ABB RobotStudio station: Project2_1.rsstnx

Station Project2 (saved by RobotStudio 25.5.11605.0)
Controller Controller1
  mechanical unit ROB_1: IRB1090_3_58__02, 6 joints, base frame (0, 0, 0) mm
Layout (positions relative to the parent item):
  - IRB1090_3_58__02 [mechanism, from %ABB.RobotStudio.Models.IRB1090%\IRB1090_3_58__01.rslib] at (0, 0, 0) mm; joint values [-0.1802, 0.1972, 0.0337, -0.0141, 1.3827, 4.496] (rad or m)
  - SOURCE AREA [graphiccomponentgroup, from Equipment\Euro Pallet.rslib] at (-200, 120, 0) mm
    - Body 1 [part, from Equipment\Euro Pallet.rslib]
  - RED_SORT_AREA [graphiccomponentgroup, from Equipment\Euro Pallet.rslib] at (-200, -920, 0) mm
    - Body 1 [part, from Equipment\Euro Pallet.rslib]
  - Source_R04 [part], size 150 x 149.2 x 50 mm
  - Source_R02 [part] at (-160, 0, 0) mm, size 150 x 149.2 x 50 mm
  - Source_R05 [part] at (-90, 150, 0) mm, size 150 x 149.2 x 50 mm
  - Source_G04 [part] at (0, 0, 50) mm, size 150 x 149.2 x 50 mm
  - Source_R03 [part] at (0, 0, 100) mm, size 150 x 149.2 x 50 mm
  - Source_G03 [part] at (0, 0, 150) mm, size 150 x 149.2 x 50 mm
  - Source_G02 [part] at (-160, 0, 50) mm, size 150 x 149.2 x 50 mm
  - Source_G01 [part] at (-160, 0, 100) mm, size 150 x 149.2 x 50 mm
  - Source_R01 [part] at (-160, 0, 150) mm, size 150 x 149.2 x 50 mm
  - Source_G07 [part] at (-90, 150, 50) mm, size 150 x 149.2 x 50 mm
  - Source_G06 [part] at (-90, 150, 100) mm, size 150 x 149.2 x 50 mm
  - Source_G05 [part] at (-90, 150, 150) mm, size 150 x 149.2 x 50 mm
  - SG_EE [smart component] at (327.71, -364.56, -73.2) mm, rotated rx 2.57 ry 0.1 rz 92.24 deg
      signals: DI To_Grasp, DO Red_Detected, DO Green_Detected
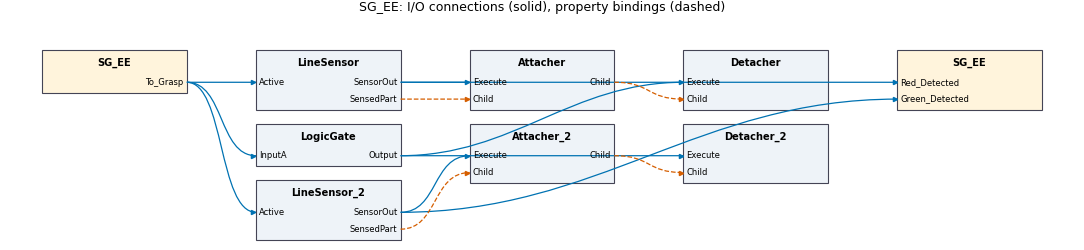
      connections:
        SG_EE.To_Grasp -> LineSensor.Active
        SG_EE.To_Grasp -> LogicGate.InputA
        LogicGate.Output -> Detacher.Execute
        LineSensor.SensorOut -> Attacher.Execute
        SG_EE.To_Grasp -> LineSensor_2.Active
        LineSensor_2.SensorOut -> Attacher_2.Execute
        LogicGate.Output -> Detacher_2.Execute
        LineSensor.SensorOut -> SG_EE.Red_Detected
        LineSensor_2.SensorOut -> SG_EE.Green_Detected
        LineSensor.SensedPart => Attacher.Child
        Attacher.Child => Detacher.Child
        LineSensor_2.SensedPart => Attacher_2.Child
        Attacher_2.Child => Detacher_2.Child
    - LogicGate [smart component, from Components\LogicGate.rslib]
        properties: Operator=NOT; Delay=0
    - LineSensor [smart component, from Components\LineSensor.rslib] at (0, 0, 50) mm
        properties: Start=[0.3 0 0.435]; End=[0.3 0 0.425]; Length=0.00999999999999995; Radius=0.0110132158590308; Tag=Tag_1; SenseMultiple=false; SensedPart=(none); SensedPoint=[0 0 0]
      - _sensorPart_ [part], size 22 x 22 x 10 mm
    - Attacher [smart component, from Components\Attacher.rslib]
        properties: Parent=EE_tool; Flange=0; Child=(none); Mount=false; Offset=[0 0 0]; Orientation=[0 0 0]
    - Detacher [smart component, from Components\Detacher.rslib]
        properties: Child=(none); KeepPosition=true
    - EE_tool [mechanism] at (299.85, 0, 553) mm, rotated rx 180 ry -0.14 rz 180 deg
        TCP EE_tool at (0, 0, -70) mm, rotated rx 180 ry 0 rz 0 deg
        links: EE
    - LineSensor_2 [smart component, from Components\LineSensor.rslib]
        properties: Start=[0.300468401861399 -2.79720985579823E-06 0.484511357513637]; End=[0.300525732933959 0.000547750941646302 0.474476736948762]; Length=0.0100498756211209; Radius=0.0108695652173913; Tag=Tag_2; SenseMultiple=false; SensedPart=(none); SensedPoint=[0 0 0]
      - _sensorPart_ [part], size 21.7 x 22.1 x 11.2 mm
    - Attacher_2 [smart component, from Components\Attacher.rslib]
        properties: Parent=EE_tool; Flange=0; Child=(none); Mount=false; Offset=[0 0 0]; Orientation=[0 0 0]
    - Detacher_2 [smart component, from Components\Detacher.rslib]
        properties: Child=(none); KeepPosition=true
Attachment: EE_tool is attached to IRB1090_3_58__02 / Link6
Attachment: SG_EE is attached to IRB1090_3_58__02 / Link6
Station logic (signal -> signal, property => property):
  Controller1.to_grasp_signal -> SG_EE.To_Grasp
  SG_EE.Red_Detected -> Controller1.red_detect
  SG_EE.Green_Detected -> Controller1.green_detect
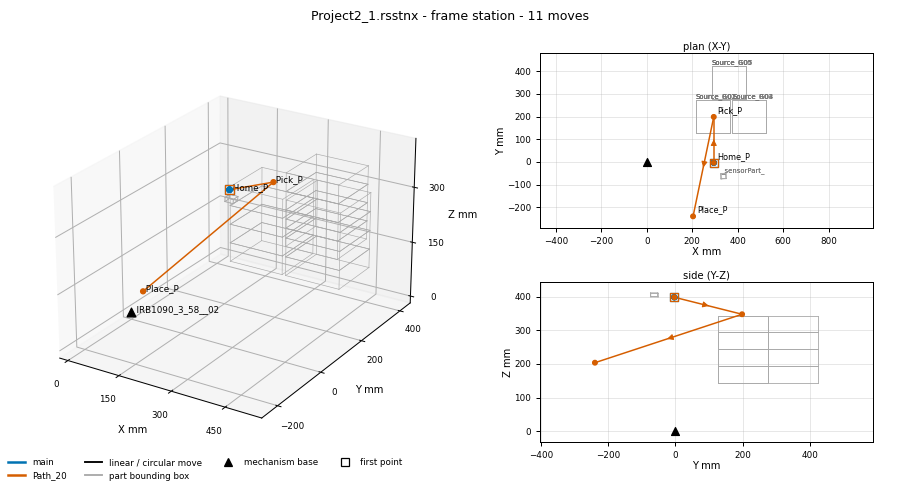
[picture p0: tool path of Project2_1.rsstnx in frame station, 11 of 26 moves have a stored position in this frame; points joined in program order, loops and branches not executed]
Targets, tools, work objects and paths stored in the station, written as RAPID:
! task T_ROB1
MODULE CalibData
  PERS tooldata EE_tool:=[TRUE,[[0,0,70],[1,0,0,0]],[1,[0,0,1],[1,0,0,0],0,0,0]];
ENDMODULE

! task T_ROB1
MODULE Module1
  CONST robtarget Pick_P:=[[294.42656998,198.457700497,347.964193384],[0.017587783,0.720617677,-0.692967877,-0.014012659],[0,0,3,0],[9E+09,9E+09,9E+09,9E+09,9E+09,9E+09]];
  CONST robtarget Home_P:=[[294.426577069,-3.238928977,398.626204981],[0.017587782,0.720617719,-0.692967834,-0.014012666],[-1,-1,2,0],[9E+09,9E+09,9E+09,9E+09,9E+09,9E+09]];
  CONST robtarget Place_P:=[[203.317190624,-239.378192774,203.819803513],[0.01758777,0.720617732,-0.692967821,-0.014012625],[-1,-1,2,0],[9E+09,9E+09,9E+09,9E+09,9E+09,9E+09]];
  CONST robtarget GreenPlace_P:=[[203.317190624,-89.378192774,203.819803513],[0.01758777,0.720617732,-0.692967821,-0.014012625],[-1,-1,2,0],[9E+09,9E+09,9E+09,9E+09,9E+09,9E+09]];
  CONST robtarget RedPlace_P:=[[203.317190624,-239.378192774,203.819803513],[0.01758777,0.720617732,-0.692967821,-0.014012625],[-1,-1,2,0],[9E+09,9E+09,9E+09,9E+09,9E+09,9E+09]];
  CONST robtarget Red_Place_P:=[[203.317190624,-239.378192774,203.819803513],[0.01758777,0.720617732,-0.692967821,-0.014012625],[-1,-1,2,0],[9E+09,9E+09,9E+09,9E+09,9E+09,9E+09]];
  CONST robtarget Green_Place_P:=[[-350,0,0],[0.01758777,0.720617732,-0.692967821,-0.014012625],[-1,-1,2,0],[9E+09,9E+09,9E+09,9E+09,9E+09,9E+09]];
  PROC main()
    MoveL Home_P,v100,fine,EE_tool\WObj:=wobj0;
    Reset To_grasp_signal;
    MoveL Offs(Pick_P,0,0,-50*i),v100,fine,EE_tool\WObj:=wobj0;
    Set To_grasp_signal;
    MoveL Home_P,v100,fine,EE_tool\WObj:=wobj0;
    MoveL Offs(Red_Place_P,
                           0,
                           0,
                           150 + 50*red_count),v50,fine,EE_tool\WObj:=wobj0;
    MoveL Offs(Red_Place_P,
                           0,
                           0,
                           50*red_count),v50,fine,EE_tool\WObj:=wobj0;
    Reset To_grasp_signal;
    MoveL Offs(Green_Place_P,
                           0,
                           0,
                           150 + 50*green_count),v50,fine,EE_tool\WObj:=wobj0;
    MoveL Offs(Green_Place_P,
                           0,
                           0,
                           50*green_count),v50,fine,EE_tool\WObj:=wobj0;
    Reset To_grasp_signal;
    MoveL Home_P,v100,fine,EE_tool\WObj:=wobj0;
    MoveL Offs(Pick_P,160,0,-50*i),v100,fine,EE_tool\WObj:=wobj0;
    Set To_grasp_signal;
    MoveL Home_P,v100,fine,EE_tool\WObj:=wobj0;
    MoveL Offs(Red_Place_P,
                           0,
                           0,
                           150 + 50*red_count),v50,fine,EE_tool\WObj:=wobj0;
    MoveL Offs(Red_Place_P,
                           0,
                           0,
                           50*red_count),v50,fine,EE_tool\WObj:=wobj0;
    Reset To_grasp_signal;
    MoveL Offs(Green_Place_P,
                           0,
                           0,
                           150 + 50*green_count),v50,fine,EE_tool\WObj:=wobj0;
    MoveL Offs(Green_Place_P,
                           0,
                           0,
                           50*green_count),v50,fine,EE_tool\WObj:=wobj0;
    Reset To_grasp_signal;
    MoveL Home_P,v100,fine,EE_tool\WObj:=wobj0;
    MoveL Offs(Pick_P,70,150,-50*i),v100,fine,EE_tool\WObj:=wobj0;
    Set To_grasp_signal;
    MoveL Home_P,v100,fine,EE_tool\WObj:=wobj0;
    MoveL Offs(Red_Place_P,
                           0,
                           0,
                           150 + 50*red_count),v50,fine,EE_tool\WObj:=wobj0;
    MoveL Offs(Red_Place_P,
                           0,
                           0,
                           50*red_count),v50,fine,EE_tool\WObj:=wobj0;
    Reset To_grasp_signal;
    MoveL Offs(Green_Place_P,
                           0,
                           0,
                           150 + 50*green_count),v50,fine,EE_tool\WObj:=wobj0;
    MoveL Offs(Green_Place_P,
                           0,
                           0,
                           50*green_count),v50,fine,EE_tool\WObj:=wobj0;
    Reset To_grasp_signal;
    MoveL Home_P,v100,fine,EE_tool\WObj:=wobj0;
    Reset To_grasp_signal;
    MoveL Home_P,v100,fine,EE_tool\WObj:=wobj0;
  ENDPROC
  PROC Path_20()
    MoveL Home_P,v1000,z100,EE_tool\WObj:=wobj0;
    MoveL Pick_P,v1000,z100,EE_tool\WObj:=wobj0;
    MoveL Place_P,v1000,z100,EE_tool\WObj:=wobj0;
  ENDPROC
ENDMODULE

